SUBAPPLICATION Button_IXA_TO_Remote_WRITE_BG_OPC (* VT-Button lesen + Remote-OPC-UA-Write an Zielmodul + VT-Hintergrundfarbe aus Remote-Subscribe (generisch, ein Kanal, fuer Ausgaenge auf Modulen ohne eigene VT-Anbindung) *)
  (* Standard: 61499-2 *)
  (* Version 1.0, 2026-08-27, franz, Meisterschulen am Ostbahnhof *)
  PACKAGE MyLib::sys;
  IMPORT isobus::UT::Q::const::IDs::ID_NULL;
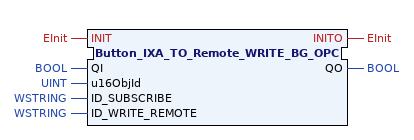
  EVENT_INPUT
    INIT : EInit; (* Initialization Request *)
  END_EVENT
  EVENT_OUTPUT
    INITO : EInit; (* Initialization Confirm *)
  END_EVENT
  VAR_INPUT
    QI : BOOL := TRUE; (* Quality Input - TRUE to enable service *)
    u16ObjId : UINT := ID_NULL; (* Object ID Button/Hintergrund (VT) *)
    ID_SUBSCRIBE : WSTRING; (* Remote-Subscribe-Adresse (Status/Farbe, ACTION=SUBSCRIBE) *)
    ID_WRITE_REMOTE : WSTRING; (* Remote-Write-Adresse zum Zielmodul (Befehl, ACTION=WRITE, CLIENT) *)
  END_VAR
  VAR_OUTPUT
    QO : BOOL; (* Quality Output - TRUE if service executed successfully *)
  END_VAR
  FBS
    Button_IXA : isobus::UT::io::Button::Button_IXA;
    AX_CLIENT_1_0 : adapter::net::AX_CLIENT_1_0;
    AX_SUBSCRIBE_1 : adapter::net::AX_SUBSCRIBE_1;
    AND_QO : iec61131::booleanOperators::AND_BOOL_4;
  END_FBS
  SUBAPPS
    GreenWhiteBackground1_AX : MyLib::sys::GreenWhiteBackground1_AX;
  END_SUBAPPS
  EVENT_CONNECTIONS
    INIT TO Button_IXA.INIT;
    Button_IXA.INITO TO AX_CLIENT_1_0.INIT;
    AX_CLIENT_1_0.INITO TO AX_SUBSCRIBE_1.INIT;
    AX_SUBSCRIBE_1.INITO TO GreenWhiteBackground1_AX.INIT;
    GreenWhiteBackground1_AX.INITO TO INITO;
    GreenWhiteBackground1_AX.INITO TO AND_QO.REQ;
  END_CONNECTIONS
  DATA_CONNECTIONS
    u16ObjId TO Button_IXA.u16ObjId;
    u16ObjId TO GreenWhiteBackground1_AX.u16ObjId;
    ID_SUBSCRIBE TO AX_SUBSCRIBE_1.ID;
    ID_WRITE_REMOTE TO AX_CLIENT_1_0.ID;
    QI TO Button_IXA.QI;
    QI TO AX_CLIENT_1_0.QI;
    QI TO AX_SUBSCRIBE_1.QI;
    Button_IXA.QO TO AND_QO.IN1;
    AX_CLIENT_1_0.QO TO AND_QO.IN2;
    AX_SUBSCRIBE_1.QO TO AND_QO.IN3;
    AND_QO.OUT TO QO;
    QI TO GreenWhiteBackground1_AX.QI;
    GreenWhiteBackground1_AX.QO TO AND_QO.IN4;
  END_CONNECTIONS
  ADAPTER_CONNECTIONS
    Button_IXA.IN TO AX_CLIENT_1_0.IN;
    AX_SUBSCRIBE_1.OUT TO GreenWhiteBackground1_AX.DI1;
  END_CONNECTIONS
END_SUBAPPLICATION
